(* IEC 61131-3 sources: codesys-to-s7/tests/fixtures/s7-to-codesys/src/POUs/S7Compat/F_ScaleX, 1 file *)

(* ---- F_ScaleX.decl.st ---- *)
// Назначение: аналог инструкции S7 SCALE_X (S7-1200/1500) для кода, сконвертированного s7conv:
//             масштабирование OUT = VALUE * (MAX - MIN) + MIN. VALUE вне 0.0…1.0 не
//             ограничивается: результат линейно продолжается за MIN и MAX (в S7 при этом
//             ENO = TRUE). При MIN >= MAX — та же формула (в S7 ENO = FALSE, значение OUT не
//             документировано — сверить с источником). Целый OUT S7 (INT, DINT) эмиттер получает
//             преобразованием REAL_TO_<тип> — округление сверить с S7. ENO не воспроизводится.
// Автор:      kr0nsch
// Версия:     0.1.0
// Документ:   docs/MAPPING.md, раздел «NORM_X и SCALE_X»
FUNCTION F_ScaleX : REAL
VAR_INPUT
    rMin : REAL;        // нижняя граница диапазона результата (MIN в S7)
    rValue : REAL;      // нормированное значение, номинально 0.0…1.0 (VALUE в S7)
    rMax : REAL;        // верхняя граница диапазона результата (MAX в S7)
END_VAR
